// TwinCAT 3 PLC project TankPLC
// ProgramVersion: 3.1.4026.27
// CompilerDefines: VISU_USEPROPERTYINFO
// libraries:
//   Tc2_Standard, * (Beckhoff Automation GmbH)
//   Tc2_System, * (Beckhoff Automation GmbH)
//   VisuSymbols, 4.5.0.0 (System)
// project tree:
//   DUTs/ E_TankFault.TcDUT, E_TankState.TcDUT, ST_TankHMI.TcDUT, E_SystemState.TcDUT
//   / GlobalTextList.TcGTLO, PlcTask.TcTTO, Visualization Manager.TcVMO (not stored)
//   GVLs/ GVL_HMI.TcGVL, GVL_IO.TcGVL
//   POUs/ FB_SystemSM.TcPOU, FB_TankControl.TcPOU, FB_TankPlantSim.TcPOU, FB_TankSM.TcPOU, MAIN.TcPOU
//   VISUs/ TankVisual.TcVIS
// real-time tasks:
//   TASK PlcTask: cycle T#10ms, priority 20, ADS port 350

CONFIGURATION TankPLC
    RESOURCE PLC ON TwinCAT3
        TASK PlcTask(INTERVAL := T#10ms, PRIORITY := 20);
        PROGRAM MAIN WITH PlcTask : MAIN;
    END_RESOURCE
END_CONFIGURATION

// ---- DUTs/E_TankFault.TcDUT
{attribute 'qualified_only'}
{attribute 'strict'}
TYPE E_TankFault :
(
    None           := 0,
    EStop          := 1,
    BusFault       := 2,
    SensorMismatch := 3,
    FillTimeout    := 4,
    DrainTimeout   := 5
) INT;
END_TYPE

// ---- DUTs/E_TankState.TcDUT
{attribute 'qualified_only'}
{attribute 'strict'}
TYPE E_TankState :
(
	Idle	:= 0,
	Filling := 10,
	Full	:= 20,
	Draining := 30,
	Empty	:= 35,
	Manual	:= 40,
	Fault	:= 99
) INT;
END_TYPE

// ---- DUTs/ST_TankHMI.TcDUT
TYPE ST_TankHMI :
STRUCT
    // ---- Commands (HMI -> PLC) ----
    bAutoMode      : BOOL;
    bStart         : BOOL;
    bStop          : BOOL;
    bReset         : BOOL;
    bPB_ValveIn    : BOOL;
    bPB_ValveOut   : BOOL;
    bPB_Pump       : BOOL;

    // ---- Status (PLC -> HMI) ----
    bLampValveIn   : BOOL;
    bLampValveOut  : BOOL;
    bLampPump      : BOOL;
    bLampHigh      : BOOL;
    bLampLow       : BOOL;
    bFaultActive   : BOOL;
    eState         : E_TankState;
    eFaultCode     : E_TankFault;
	
	rLevel         : REAL; 
END_STRUCT
END_TYPE

// ---- DUTs/E_SystemState.TcDUT
{attribute 'qualified_only'}
{attribute 'strict'}
TYPE E_SystemState :
(
	Start 	:= 0,
	Stop 	:= 1,
	Reset	:= 2,
	Fault	:= 99
) INT;
END_TYPE

// ---- GVLs/GVL_HMI.TcGVL
{attribute 'qualified_only'}
VAR_GLOBAL
    Tank1 : ST_TankHMI;
END_VAR

// ---- GVLs/GVL_IO.TcGVL
{attribute 'qualified_only'}
VAR_GLOBAL
	// IN
	bSensHigh_RAW	AT %I* : BOOL;
	bSensLow_RAW	AT %I* : BOOL;
	bEStop_RAW		AT %I* : BOOL;
	
	// OUT
	bValveIn		AT %Q* : BOOL;
	bValveOut		AT %Q* : BOOL;
	bPump			AT %Q* : BOOL;
END_VAR

// ---- POUs/MAIN.TcPOU
PROGRAM MAIN
VAR
	// Create instance of FB
	Tank1SM : FB_TankSM;
	
	// Internal Bools to handle I/O inputs
	bEStopPressed 	: BOOL; // TRUE = PRESSED (inverted from raw)
	bSensHIGH		: BOOL;
	bSensLOW		: BOOL;
	bBusOK			: BOOL := TRUE; // Practical IRL but unused in this simulation.
	
	// Timers
	tTankfillTimeout	: TIME := T#120S; 
	
	// FB Outputs
	bValveInCMD		: BOOL;
	bValveOutCMD	: BOOL;
	bPumpCMD		: BOOL;
	bTankFault		: BOOL;
	bAutoMode		: BOOL;
	
	eTankState		: E_TankState;
	eTankFaultCode  : E_TankFault;
	eSystemState	: E_SystemState;
	
	// Plant-level
	bOutputsDisabled : BOOL; // practical IRL for maitinence lockout, but unused in this simulation
	fbHeartbeat		: TON;
	bHeartbeat		: BOOL;
	
	// ---- Simulation ----
    fbSim            : FB_TankPlantSim;
    bSimMode         : BOOL := TRUE;     // TRUE = no hardware, use fbSim
    bSimEStop        : BOOL;             // HMI toggle: simulated e-stop pressed
    bSimBusOK        : BOOL := TRUE;     // HMI toggle: simulated bus health
	// Final outputs after plant-level overrides 
    bOutValveIn      : BOOL;
    bOutValveOut     : BOOL;
    bOutPump         : BOOL;


END_VAR

// Main will primarily call function blocks in order

// Pull in I/O Inputs from GVL (or in this case, the SIM)
bSensHIGH     := fbSim.bSensHIGH;
bSensLOW      := fbSim.bSensLOW;
bEStopPressed := bSimEStop;
bAutoMode     := GVL_HMI.Tank1.bAutoMode; 
(* This is what it would look like as GVL *)(*    
bEStopPressed := NOT GVL_IO.bEStop_RAW; 
bSensHIGH     := GVL_IO.bSensHigh_RAW;    
bSensLOW      := GVL_IO.bSensLow_RAW;
*)


// HMI COMMAND HANDLING
// This program was designed under the assumption that this MAIN may manage more than one tank.
// As such, most of the IO reaction is handled by the FB's, and results passed in the next section.

// FB CALL sysSM -> tankSM -> pumpSM -> simSM
Tank1SM(
	// These go INTO the FB :=
	bSensHIGH	:= bSensHIGH,
	bSensLOW	:= bSensLOW,
	eSystemState := eSystemState,
	
	// These come OUT of the FB =>
	eTankState => eTankState,
	bOutValveIn	=> bValveInCMD,
	bOutValveOut => bValveOutCMD,
	bOutPump => bPumpCMD,
	// VAR_IN_OUT
	bAutoMode	:= bAutoMode
);

// OUTPUT MAPING
// Plant-level overrides such as E-Stop presses, bus fault, etc. 
// For this exercise, it's not simulated but still here.
IF bOutputsDisabled OR NOT bBusOK OR bEStopPressed THEN // if something wrong, soft stop
    bOutValveIn  := FALSE;
    bOutValveOut := FALSE;
    bOutPump     := FALSE;
ELSE 
    bOutValveIn  := bValveInCMD;
    bOutValveOut := bValveOutCMD;
    bOutPump     := bPumpCMD;
END_IF;

IF bSimMode THEN
    fbSim(
        bValveIn  := bOutValveIn,
        bValveOut := bOutValveOut,
        bPump     := bOutPump,
        tCycle    := T#10MS             
    );
    GVL_HMI.Tank1.rLevel := fbSim.rLevel;

    GVL_IO.bValveIn  := FALSE;          
    GVL_IO.bValveOut := FALSE;
    GVL_IO.bPump     := FALSE;
ELSE
    GVL_IO.bValveIn  := bOutValveIn;
    GVL_IO.bValveOut := bOutValveOut;
    GVL_IO.bPump     := bOutPump;
END_IF;


// STATUS AND DIAGNOSTICS
// Things like heartbeat, warning flags, etc.
fbHeartbeat(IN := NOT fbHeartbeat.Q, PT := T#500MS);
IF fbHeartbeat.Q THEN
    bHeartbeat := NOT bHeartbeat;
END_IF;

END_PROGRAM

// ---- POUs/FB_TankSM.TcPOU
FUNCTION_BLOCK FB_TankSM
VAR_INPUT
	bSensHIGH, bSensLOW	: BOOL;
	bFaultClear			: BOOL;
	bBusOK				: BOOL;
	bTankFault				: BOOL;
	
	eTankFaultCode		: E_TankFault;
	eSystemState		: E_SystemState;
	
	// passed in from TankCrontrol to go to Main
	bValveIn    : BOOL;
    bValveOut   : BOOL;
    bPump       : BOOL;
END_VAR
VAR_OUTPUT
	eTankState				: E_TankState;
	
	// pass from TankControl to Main
	bOutValveIn				: BOOL;
	bOutValveOut			: BOOL;
	bOutPump				: BOOL;
END_VAR
VAR_IN_OUT
	bAutoMode			: BOOL;
END_VAR
VAR
	TankCTRL	: FB_TankControl;
	
    tonEmptyDelay     : TON;
	tonPumpStartDelay : TON;
	tonStayFull		  : TON;
	tEmptyDelay       : TIME := T#2S;
	tPumpStartDelay   : TIME := T#3S;
	tStayFullTime	  : TIME := T#3S;
	
	bcmdOpenValveIn 		: BOOL;
	bcmdOpenValveOut		: BOOL;
	bcmdPumpOn				: BOOL;
END_VAR

// State Machine for the Tank

IF NOT bAutoMode THEN
	eTankState := 40;
END_IF
IF eSystemState = 99 OR bTankFault THEN
	eTankState := 99;
END_IF

tonEmptyDelay(IN := (eTankState = 35), PT := tEmptyDelay);
tonPumpStartDelay(IN := (eTankState = 10), PT := tPumpStartDelay);
tonStayFull(IN := (eTankState = 20), PT := tStayFullTime);

CASE eTankState OF
	0://IDLE 
		IF NOT bSensHIGH AND NOT bSensLOW THEN // Empty
			eTankState := 35;
		ELSIF bSensLOW THEN //If between sensors then go to filling
			eTankState := 10;
		ELSE // if high then drain
			eTankState := 30;
		END_IF
	10://FILLING
	bcmdOpenValveIn := TRUE;
		bcmdPumpOn := TRUE;
		 IF tonPumpStartDelay.Q AND bSensHIGH THEN
			bcmdOpenValveIn := FALSE; // close in valve; full
			eTankState := 20;
		END_IF
	20://FULL
		IF tonStayFull.Q THEN
			eTankState := 30; // drain after 3s
		ELSIF NOT bSensHIGH THEN // if no longer high then trigger into idle
			bcmdPumpOn := FALSE;
			eTankState := 0;
		END_IF
	30: // DRAINING
		bcmdOpenValveOut := TRUE;
        IF NOT bSensLOW THEN
            bcmdOpenValveOut := FALSE;
            eTankState := 35;
        END_IF
    35: // EMPTY - hold 2 s before starting to fill
        IF tonEmptyDelay.Q THEN
            eTankState := 10;
        END_IF
	40://MANUAL
		IF bAutoMode THEN
			eTankState := 0;
		END_IF
	99://FAULT
		bcmdPumpOn := FALSE;
		IF bFaultClear THEN
			eTankState := 0;
		END_IF
END_CASE

TankCTRL(
    // Commands from the state machine
    cmdOpenValveIn  := bcmdOpenValveIn,
    cmdOpenValveOut := bcmdOpenValveOut,
    cmdPumpOn       := bcmdPumpOn,
    bAutoMode       := bAutoMode,

    // Status
    bFault          => bTankFault,
    eFaultCode      => eTankFaultCode,
    bBusOK          => bBusOK,

    // Final outputs, passed straight through to MAIN
    bValveIn        => bOutValveIn,
    bValveOut       => bOutValveOut,
    bPump           => bOutPump
);

END_FUNCTION_BLOCK

// ---- POUs/FB_TankControl.TcPOU
FUNCTION_BLOCK FB_TankControl
VAR_INPUT
	// COMMANDS SENT BY SM
	cmdOpenValveIn 		: BOOL;
	cmdOpenValveOut		: BOOL;
	cmdPumpOn			: BOOL;
	
	bAutoMode			: BOOL;
END_VAR
VAR_OUTPUT
	bFault				: BOOL;
	eFaultCode			: E_TankFault;
	bBusOK				: BOOL; //EtherCAT
	
	bValveIn    : BOOL;
    bValveOut   : BOOL;
    bPump       : BOOL;
END_VAR
VAR_IN_OUT
END_VAR
VAR
		HMI					: ST_TankHMI;
END_VAR

// Does the physical switching for FB_TankSM

IF bAutoMode THEN
	IF cmdOpenValveIn THEN
		bValveIn := TRUE;
	ELSE
		bValveIn := FALSE;
	END_IF
	IF cmdOpenValveOut THEN
		bValveOut := TRUE;
	ELSE
		bValveOut := FALSE;
	END_IF
	IF cmdPumpOn THEN
		bPump := TRUE;
	ELSE
		bPump := FALSE;
	END_IF
ELSE
	Manual();
END_IF

METHOD Manual : BOOL
VAR_INPUT
END_VAR
// When running a tank manually, simply pass raw HMI inputs
// just push raw inputs
bValveIn  := GVL_HMI.Tank1.bPB_ValveIn;
bValveOut := GVL_HMI.Tank1.bPB_ValveOut;
bPump     := GVL_HMI.Tank1.bPB_Pump;
END_METHOD

END_FUNCTION_BLOCK

// ---- POUs/FB_TankPlantSim.TcPOU
FUNCTION_BLOCK FB_TankPlantSim
VAR_INPUT
    bValveIn          : BOOL;
    bValveOut         : BOOL;
    bPump             : BOOL;

    tCycle            : TIME := T#10MS;   // must match the PlcTask cycle time

    rFillRate         : REAL := 8.0;      // % per second, pump running AND inlet open
    rDrainRate        : REAL := 6.0;      // % per second, outlet open (gravity)
    rHighSP           : REAL := 85.0;     // level where SENS HIGH goes wet
    rLowSP            : REAL := 15.0;     // level where SENS LOW goes wet

    // Fault injection: set from the HMI, NOT passed in the call from MAIN
    bFailHighDry      : BOOL;             // high sensor stuck reading dry
    bFailLowDry       : BOOL;             // low sensor stuck reading dry
    bResetLevel       : BOOL;             // empty the tank
END_VAR
VAR_OUTPUT
    rLevel            : REAL;             // 0..100 %
    bSensHIGH         : BOOL;
    bSensLOW          : BOOL;
END_VAR
VAR
    rDt               : REAL;             // cycle time in seconds
END_VAR

// Simulation FB

rDt := TIME_TO_REAL(tCycle) / 1000.0;     // TIME_TO_REAL gives milliseconds

IF bResetLevel THEN
    rLevel := 0.0;
END_IF;

// Inflow: the pump feeds the inlet line. Liquid only moves if the inlet
// valve is open too (pump against a closed valve = dead-head, no flow).
IF bPump AND bValveIn THEN
    rLevel := rLevel + rFillRate * rDt;
END_IF;

// Outflow: gravity drain through the outlet valve
IF bValveOut THEN
    rLevel := rLevel - rDrainRate * rDt;
END_IF;

rLevel := LIMIT(0.0, rLevel, 100.0);

// Sensors, with optional injected failures
bSensHIGH := (rLevel >= rHighSP) AND NOT bFailHighDry;
bSensLOW  := (rLevel >= rLowSP)  AND NOT bFailLowDry;

END_FUNCTION_BLOCK

// ---- POUs/FB_SystemSM.TcPOU
FUNCTION_BLOCK FB_SystemSM
VAR_INPUT
END_VAR
VAR_OUTPUT
END_VAR
VAR
END_VAR

// Edge-Detect Commands
// MOVE ME!!
//_TrigStart(CLK := HMI.bStart);
//_TrigStop(CLK := HMI.bStop);
//_TrigReset(CLK := HMI.bReset);

END_FUNCTION_BLOCK

// ---- GlobalTextList.TcGTLO
TEXTLIST GlobalTextList
  151 = '%s'
  168 = 'Auto'
  12 = 'Auto/Manual'
  840 = 'Fault'
  497 = 'In Valve'
  392 = 'Label'
  586 = 'Out Valve'
  620 = 'Pump'
  33 = 'Reset'
  972 = 'Start'
  729 = 'Start/Stop/Reset'
  506 = 'State'
  8 = 'Stop'
END_TEXTLIST

// ---- VISUs/TankVisual.TcVIS
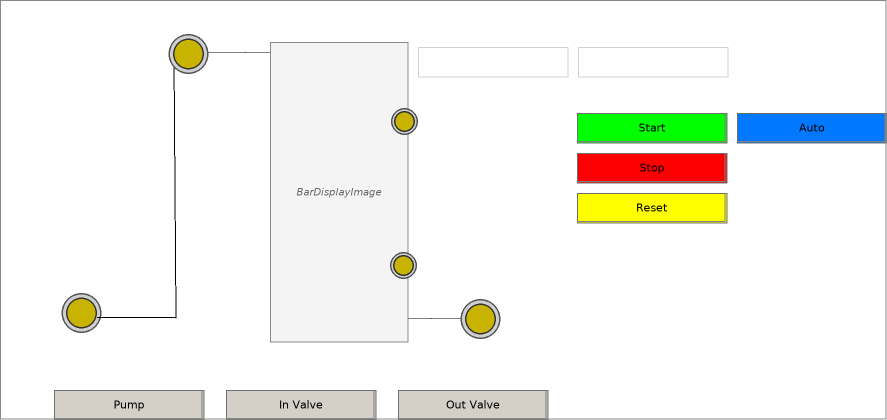
VISUALIZATION TankVisual  // 887x420
    Line (474,319) (389,318)
    Line (288,53) (203,52)
    Rectangle (270,42 138x300)
    BarDisplayImage (270,42 138x300), value: GVL_HMI.Tank1.rLevel, style: BarDisplayImage-Gray, scale format: %.1f, scale 0..100
    Lamp1 (453,296 55x46), variable: GVL_HMI.Tank1.bPB_ValveOut, style: Lamp-Lamp1-Yellow
    Lamp1 (54,290 55x46), variable: GVL_HMI.Tank1.bPB_Pump, style: Lamp-Lamp1-Yellow
    Lamp1 (389,106 31x31), variable: MAIN.bSensHIGH, style: Lamp-Lamp1-Yellow
    Lamp1 (388,250 31x31), variable: MAIN.bSensLOW, style: Lamp-Lamp1-Yellow
    Button (577,113 150x30), "Start", pressed state: GVL_HMI.Tank1.bStart
    Button (737,113 150x30), "Auto", pressed state: GVL_HMI.Tank1.bAutoMode
        toggle GVL_HMI.Tank1.bAutoMode p2164770859=TRUE
    Button (54,390 150x30), "Pump", input disabled if: GVL_HMI.Tank1.bAutoMode
        tap GVL_HMI.Tank1.bPB_Pump
        toggle GVL_HMI.Tank1.bPB_Pump
    Button (226,390 150x30), "In Valve", input disabled if: GVL_HMI.Tank1.bAutoMode
        toggle GVL_HMI.Tank1.bPB_ValveIn
    Button (398,390 150x30), "Out Valve", input disabled if: GVL_HMI.Tank1.bAutoMode
        toggle GVL_HMI.Tank1.bPB_ValveOut
    Line (97,317) (176,317)
    Line (176,318) (174,58)
    Lamp1 (161,31 55x46), variable: GVL_HMI.Tank1.bPB_ValveIn, style: Lamp-Lamp1-Yellow
    Button (577,193 150x30), "Reset", pressed state: GVL_HMI.Tank1.bReset
    Button (577,153 150x30), "Stop", pressed state: GVL_HMI.Tank1.bStop
    Textfield (418,47 150x30), text variable: GVL_HMI.Tank1.eState
    Textfield (578,47 150x30), text variable: GVL_HMI.Tank1.eState
END_VISUALIZATION
